ADAPTER control_IMC (* Adapter Interface *)
  (* Standard: 61499-1 *)
  (* Version 0.0, 10/23/2026, macie, Schneider Electric *)
  PACKAGE Main;
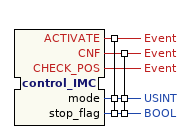
  EVENT_OUTPUT
    ACTIVATE WITH mode, stop_flag; (* Indication from Plug *)
    CNF WITH mode, stop_flag; (* Confirmation from Plug *)
    CHECK_POS;
  END_EVENT
  VAR_OUTPUT
    mode : USINT; (* Confirmation Data from Plug *)
    stop_flag : BOOL; (* Indication Data from Plug *)
  END_VAR
  SERVICE SOCKET/PLUG
    SEQUENCE request_confirm
      SOCKET.REQ(REQD) -> PLUG.REQ(REQD);
      PLUG.CNF(mode) -> SOCKET.CNF(mode);
    END_SEQUENCE
    SEQUENCE indication_response
      PLUG.ACTIVATE(stop_flag) -> SOCKET.ACTIVATE(stop_flag);
      SOCKET.RSP(RSPD) -> PLUG.RSP(RSPD);
    END_SEQUENCE
  END_SERVICE
END_ADAPTER
